(* IEC 61131-3 sources: plc-st-coding-agent/progress/v13_r4/references, 2 files *)

(* ---- self-hard-02.reference.st ---- *)
FUNCTION_BLOCK FB
VAR_INPUT
    startBtn : BOOL;
    abortBtn : BOOL;
    setpoint : REAL;
    pv : REAL;
    maxDuration : INT;
END_VAR
VAR_OUTPUT
    elapsed : INT;
    phase : INT;
    timeout : BOOL;
END_VAR
VAR
    startEdgeInputPrev : BOOL;
    startEdge : BOOL;
END_VAR
startEdge := startBtn AND NOT startEdgeInputPrev;
startEdgeInputPrev := startBtn;
IF abortBtn THEN
    phase := 9;
ELSIF startEdge THEN
    phase := 1;
    elapsed := 0;
    timeout := FALSE;
ELSIF phase = 1 OR phase = 2 THEN
    elapsed := elapsed + 1;
    IF elapsed >= maxDuration THEN
        timeout := TRUE;
        phase := 3;
    ELSIF phase = 1 AND pv >= setpoint THEN
        phase := 2;
    END_IF
END_IF
END_FUNCTION_BLOCK

(* ---- self-hard-04.reference.st ---- *)
FUNCTION_BLOCK FB
VAR_INPUT
    demand : INT;
    runHours : ARRAY[1..5] OF LINT;
    rotated : BOOL;
END_VAR
VAR_OUTPUT
    leadPump : INT;
    lagPump : INT;
    runningCount : INT;
END_VAR
VAR
    i : INT;
    j : INT;
    tmp : INT;
    need : INT;
    pickLag : BOOL;
    order : ARRAY[1..5] OF INT;
END_VAR
need := LIMIT(0, demand, 5);
FOR i := 1 TO 5 DO order[i] := i; END_FOR
FOR i := 1 TO 4 DO
    FOR j := i + 1 TO 5 DO
        IF (runHours[order[j]] < runHours[order[i]]) OR
           ((runHours[order[j]] = runHours[order[i]]) AND (order[j] < order[i])) THEN
            tmp := order[i]; order[i] := order[j]; order[j] := tmp;
        END_IF
    END_FOR
END_FOR
runningCount := need;
IF need = 0 THEN
    leadPump := 0; lagPump := 0;
ELSE
    pickLag := FALSE;
    IF leadPump = 0 THEN
        leadPump := order[1]; pickLag := TRUE;
    ELSIF rotated THEN
        IF runHours[leadPump] - runHours[order[1]] > 50 THEN
            leadPump := order[1]; pickLag := TRUE;
        END_IF
    END_IF
    IF need = 1 THEN
        lagPump := 0;
    ELSIF pickLag OR lagPump = 0 THEN
        IF order[1] <> leadPump THEN lagPump := order[1];
        ELSE lagPump := order[2]; END_IF
    END_IF
END_IF
END_FUNCTION_BLOCK
